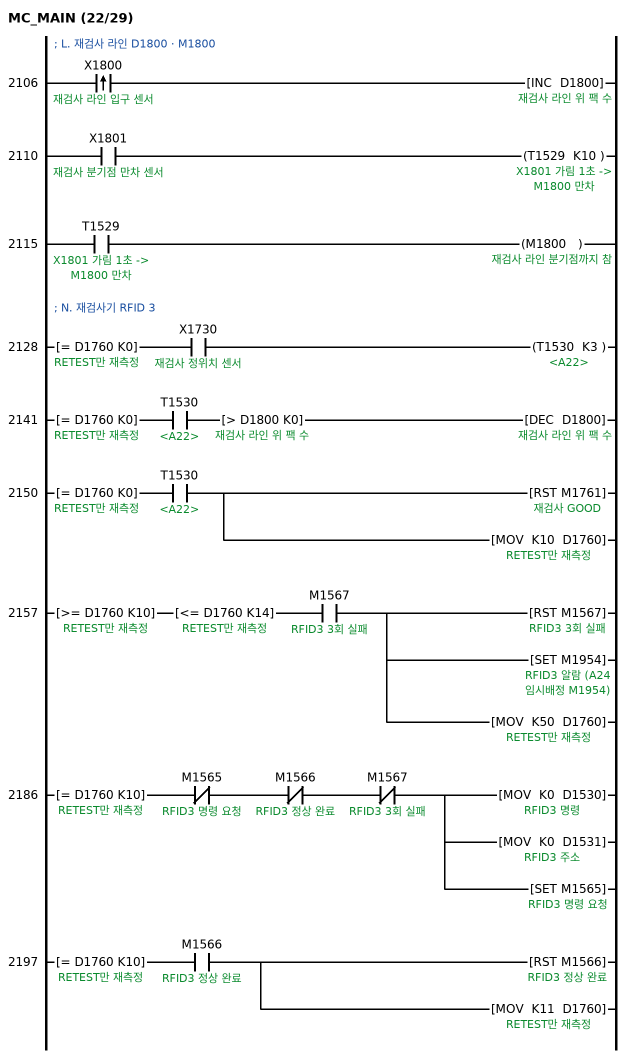
[picture p24: ladder of MC_MAIN, rungs at steps 2106 to 2197]
; L. 재검사 라인 D1800 · M1800
2106  LDP     X1800  ; 재검사 라인 입구 센서
      INC     D1800  ; 재검사 라인 위 팩 수
2110  LD      X1801  ; 재검사 분기점 만차 센서
      OUT     T1529 K10  ; X1801 가림 1초 -> M1800 만차
2115  LD      T1529  ; X1801 가림 1초 -> M1800 만차
      OUT     M1800  ; 재검사 라인 분기점까지 참
; N. 재검사기 RFID 3
2128  LD=     D1760 K0  ; RETEST만 재측정
      AND     X1730  ; 재검사 정위치 센서
      OUT     T1530 K3  ; <A22>
        [note] <A22>
2141  LD=     D1760 K0  ; RETEST만 재측정
      AND     T1530  ; <A22>
      AND>    D1800 K0  ; 재검사 라인 위 팩 수
      DEC     D1800
2150  LD=     D1760 K0  ; RETEST만 재측정
      AND     T1530  ; <A22>
      RST     M1761  ; 재검사 GOOD
      MOV     K10 D1760
2157  LD>=    D1760 K10  ; RETEST만 재측정
      AND<=   D1760 K14  ; RETEST만 재측정
      AND     M1567  ; RFID3 3회 실패
      RST     M1567  ; RFID3 3회 실패
      SET     M1954  ; RFID3 알람 (A24 임시배정 M1954)
        [note] RFID3 알람 (A24 임시배정 M1954)
      MOV     K50 D1760
2186  LD=     D1760 K10  ; RETEST만 재측정
      ANI     M1565  ; RFID3 명령 요청
      ANI     M1566  ; RFID3 정상 완료
      ANI     M1567  ; RFID3 3회 실패
      MOV     K0 D1530  ; RFID3 명령
      MOV     K0 D1531  ; RFID3 주소
      SET     M1565  ; RFID3 명령 요청
2197  LD=     D1760 K10  ; RETEST만 재측정
      AND     M1566  ; RFID3 정상 완료
      RST     M1566  ; RFID3 정상 완료
      MOV     K11 D1760
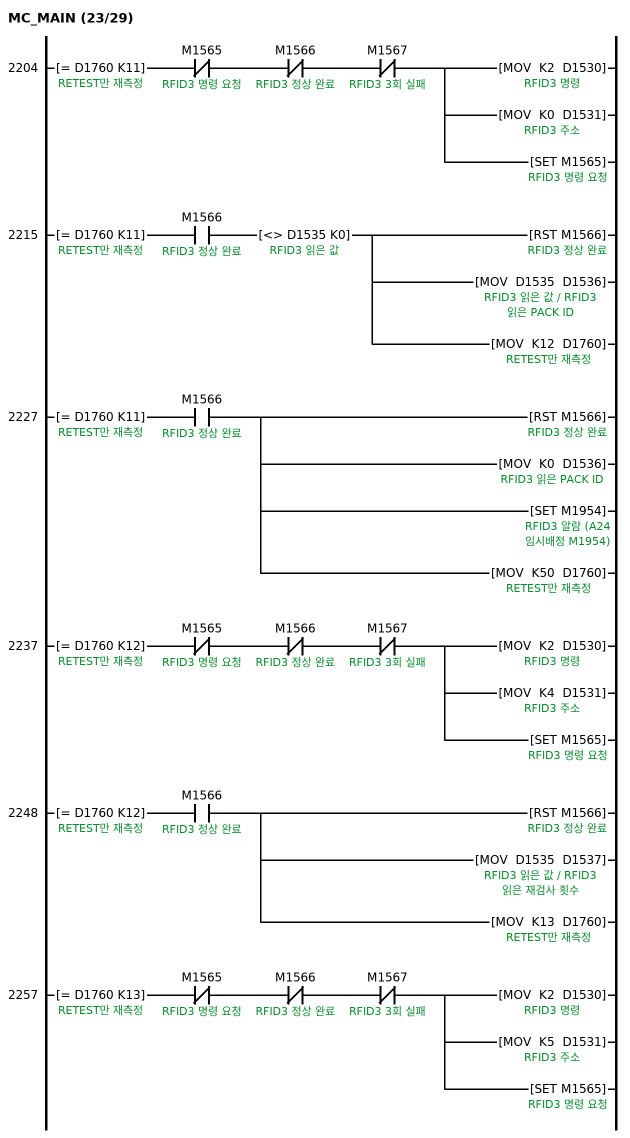
2204  LD=     D1760 K11  ; RETEST만 재측정
      ANI     M1565  ; RFID3 명령 요청
      ANI     M1566  ; RFID3 정상 완료
      ANI     M1567  ; RFID3 3회 실패
      MOV     K2 D1530
      MOV     K0 D1531
      SET     M1565  ; RFID3 명령 요청
2215  LD=     D1760 K11  ; RETEST만 재측정
      AND     M1566  ; RFID3 정상 완료
      AND<>   D1535 K0  ; RFID3 읽은 값
      RST     M1566  ; RFID3 정상 완료
      MOV     D1535 D1536  ; RFID3 읽은 PACK ID
      MOV     K12 D1760
2227  LD=     D1760 K11  ; RETEST만 재측정
      AND     M1566  ; RFID3 정상 완료
      RST     M1566  ; RFID3 정상 완료
      MOV     K0 D1536
      SET     M1954  ; RFID3 알람 (A24 임시배정 M1954)
      MOV     K50 D1760
2237  LD=     D1760 K12  ; RETEST만 재측정
      ANI     M1565  ; RFID3 명령 요청
      ANI     M1566  ; RFID3 정상 완료
      ANI     M1567  ; RFID3 3회 실패
      MOV     K2 D1530
      MOV     K4 D1531
      SET     M1565  ; RFID3 명령 요청
2248  LD=     D1760 K12  ; RETEST만 재측정
      AND     M1566  ; RFID3 정상 완료
      RST     M1566  ; RFID3 정상 완료
      MOV     D1535 D1537  ; RFID3 읽은 재검사 횟수
      MOV     K13 D1760
2257  LD=     D1760 K13  ; RETEST만 재측정
      ANI     M1565  ; RFID3 명령 요청
      ANI     M1566  ; RFID3 정상 완료
      ANI     M1567  ; RFID3 3회 실패
      MOV     K2 D1530
      MOV     K5 D1531
      SET     M1565  ; RFID3 명령 요청
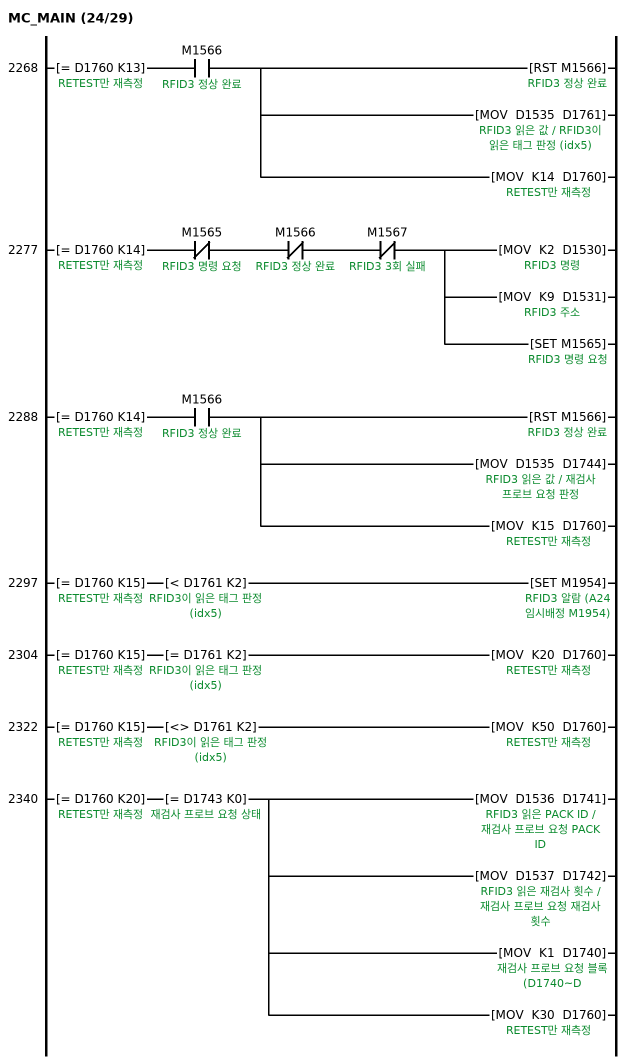
2268  LD=     D1760 K13  ; RETEST만 재측정
      AND     M1566  ; RFID3 정상 완료
      RST     M1566  ; RFID3 정상 완료
      MOV     D1535 D1761  ; RFID3이 읽은 태그 판정 (idx5)
      MOV     K14 D1760
2277  LD=     D1760 K14  ; RETEST만 재측정
      ANI     M1565  ; RFID3 명령 요청
      ANI     M1566  ; RFID3 정상 완료
      ANI     M1567  ; RFID3 3회 실패
      MOV     K2 D1530
      MOV     K9 D1531
      SET     M1565  ; RFID3 명령 요청
2288  LD=     D1760 K14  ; RETEST만 재측정
      AND     M1566  ; RFID3 정상 완료
      RST     M1566  ; RFID3 정상 완료
      MOV     D1535 D1744  ; 재검사 프로브 요청 판정
      MOV     K15 D1760
2297  LD=     D1760 K15  ; RETEST만 재측정
      AND<    D1761 K2  ; RFID3이 읽은 태그 판정 (idx5)
      SET     M1954  ; RFID3 알람 (A24 임시배정 M1954)
2304  LD=     D1760 K15  ; RETEST만 재측정
      AND=    D1761 K2  ; RFID3이 읽은 태그 판정 (idx5)
      MOV     K20 D1760
        [note] RETEST만 재측정
2322  LD=     D1760 K15  ; RETEST만 재측정
      AND<>   D1761 K2  ; RFID3이 읽은 태그 판정 (idx5)
      MOV     K50 D1760
        [note] 메인 NG -> 통과
2340  LD=     D1760 K20  ; RETEST만 재측정
      AND=    D1743 K0  ; 재검사 프로브 요청 상태
      MOV     D1536 D1741  ; 재검사 프로브 요청 PACK ID
      MOV     D1537 D1742  ; 재검사 프로브 요청 재검사 횟수
      MOV     K1 D1740  ; 재검사 프로브 요청 블록 (D1740~D
      MOV     K30 D1760
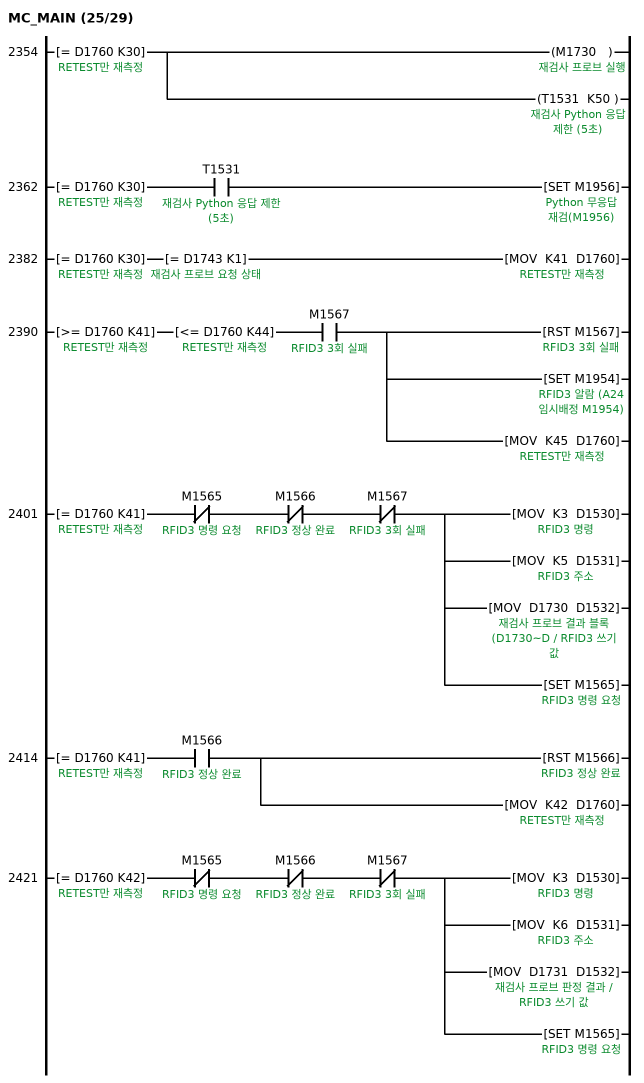
2354  LD=     D1760 K30  ; RETEST만 재측정
      OUT     M1730  ; 재검사 프로브 실행
      OUT     T1531 K50  ; 재검사 Python 응답 제한 (5초)
2362  LD=     D1760 K30  ; RETEST만 재측정
      AND     T1531  ; 재검사 Python 응답 제한 (5초)
      SET     M1956  ; Python 무응답 재검(M1956)
        [note] Python 무응답 재검(M1956)
2382  LD=     D1760 K30  ; RETEST만 재측정
      AND=    D1743 K1  ; 재검사 프로브 요청 상태
      MOV     K41 D1760
2390  LD>=    D1760 K41  ; RETEST만 재측정
      AND<=   D1760 K44  ; RETEST만 재측정
      AND     M1567  ; RFID3 3회 실패
      RST     M1567  ; RFID3 3회 실패
      SET     M1954  ; RFID3 알람 (A24 임시배정 M1954)
      MOV     K45 D1760
2401  LD=     D1760 K41  ; RETEST만 재측정
      ANI     M1565  ; RFID3 명령 요청
      ANI     M1566  ; RFID3 정상 완료
      ANI     M1567  ; RFID3 3회 실패
      MOV     K3 D1530
      MOV     K5 D1531
      MOV     D1730 D1532  ; 재검사 프로브 결과 블록 (D1730~D / RFID3 쓰기 값
      SET     M1565  ; RFID3 명령 요청
2414  LD=     D1760 K41  ; RETEST만 재측정
      AND     M1566  ; RFID3 정상 완료
      RST     M1566  ; RFID3 정상 완료
      MOV     K42 D1760
2421  LD=     D1760 K42  ; RETEST만 재측정
      ANI     M1565  ; RFID3 명령 요청
      ANI     M1566  ; RFID3 정상 완료
      ANI     M1567  ; RFID3 3회 실패
      MOV     K3 D1530
      MOV     K6 D1531
      MOV     D1731 D1532  ; 재검사 프로브 판정 결과
      SET     M1565  ; RFID3 명령 요청
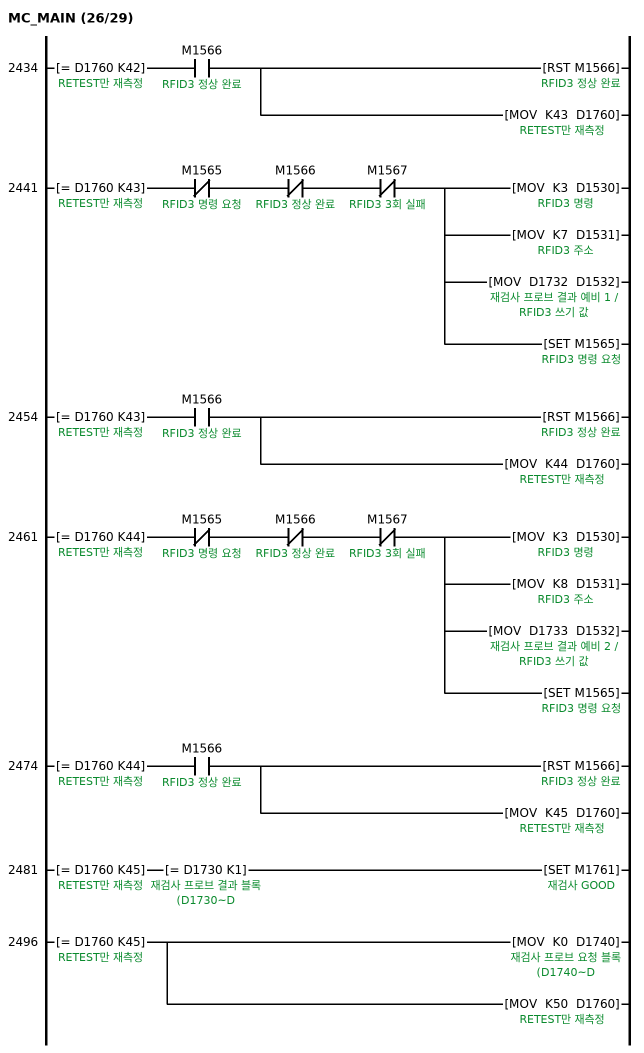
2434  LD=     D1760 K42  ; RETEST만 재측정
      AND     M1566  ; RFID3 정상 완료
      RST     M1566  ; RFID3 정상 완료
      MOV     K43 D1760
2441  LD=     D1760 K43  ; RETEST만 재측정
      ANI     M1565  ; RFID3 명령 요청
      ANI     M1566  ; RFID3 정상 완료
      ANI     M1567  ; RFID3 3회 실패
      MOV     K3 D1530
      MOV     K7 D1531
      MOV     D1732 D1532  ; 재검사 프로브 결과 예비 1
      SET     M1565  ; RFID3 명령 요청
2454  LD=     D1760 K43  ; RETEST만 재측정
      AND     M1566  ; RFID3 정상 완료
      RST     M1566  ; RFID3 정상 완료
      MOV     K44 D1760
2461  LD=     D1760 K44  ; RETEST만 재측정
      ANI     M1565  ; RFID3 명령 요청
      ANI     M1566  ; RFID3 정상 완료
      ANI     M1567  ; RFID3 3회 실패
      MOV     K3 D1530
      MOV     K8 D1531
      MOV     D1733 D1532  ; 재검사 프로브 결과 예비 2
      SET     M1565  ; RFID3 명령 요청
2474  LD=     D1760 K44  ; RETEST만 재측정
      AND     M1566  ; RFID3 정상 완료
      RST     M1566  ; RFID3 정상 완료
      MOV     K45 D1760
2481  LD=     D1760 K45  ; RETEST만 재측정
      AND=    D1730 K1  ; 재검사 프로브 결과 블록 (D1730~D
      SET     M1761  ; 재검사 GOOD
        [note] 재검사 GOOD
2496  LD=     D1760 K45  ; RETEST만 재측정
      MOV     K0 D1740
      MOV     K50 D1760
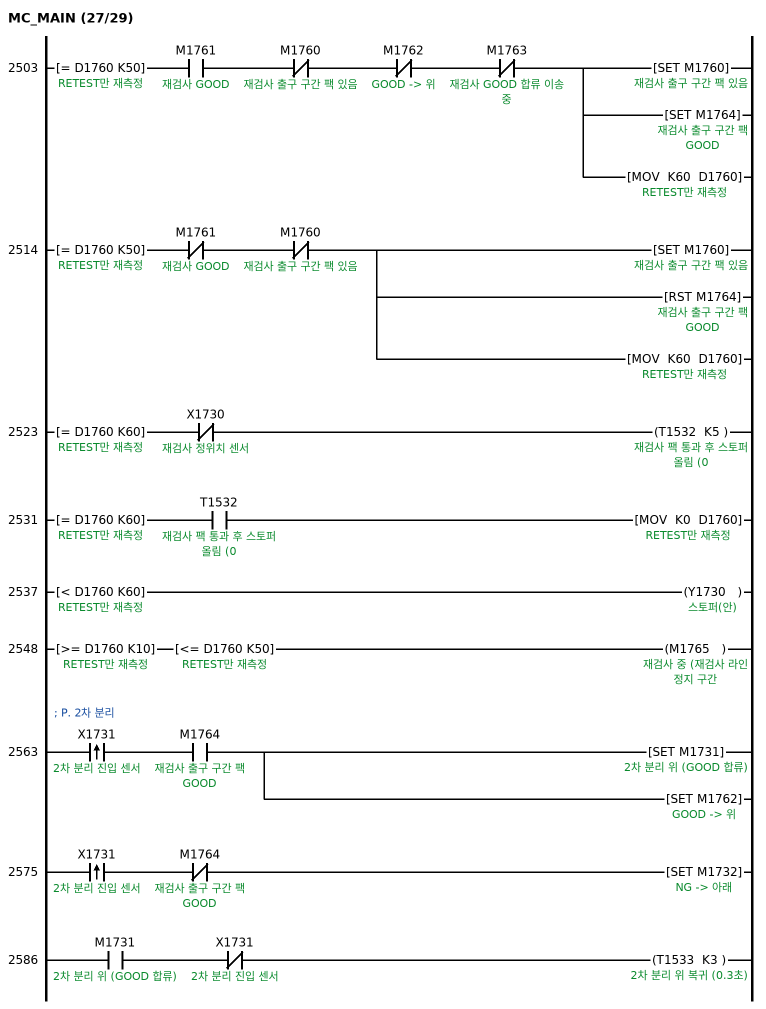
2503  LD=     D1760 K50  ; RETEST만 재측정
      AND     M1761  ; 재검사 GOOD
      ANI     M1760  ; 재검사 출구 구간 팩 있음
      ANI     M1762  ; GOOD -> 위
      ANI     M1763  ; 재검사 GOOD 합류 이송 중
      SET     M1760  ; 재검사 출구 구간 팩 있음
      SET     M1764  ; 재검사 출구 구간 팩 GOOD
      MOV     K60 D1760
2514  LD=     D1760 K50  ; RETEST만 재측정
      ANI     M1761  ; 재검사 GOOD
      ANI     M1760  ; 재검사 출구 구간 팩 있음
      SET     M1760  ; 재검사 출구 구간 팩 있음
      RST     M1764  ; 재검사 출구 구간 팩 GOOD
      MOV     K60 D1760
2523  LD=     D1760 K60  ; RETEST만 재측정
      ANI     X1730  ; 재검사 정위치 센서
      OUT     T1532 K5  ; 재검사 팩 통과 후 스토퍼 올림 (0
2531  LD=     D1760 K60  ; RETEST만 재측정
      AND     T1532  ; 재검사 팩 통과 후 스토퍼 올림 (0
      MOV     K0 D1760
2537  LD<     D1760 K60  ; RETEST만 재측정
      OUT     Y1730  ; 스토퍼(안)
        [note] 스토퍼(안)
2548  LD>=    D1760 K10  ; RETEST만 재측정
      AND<=   D1760 K50  ; RETEST만 재측정
      OUT     M1765  ; 재검사 중 (재검사 라인 정지 구간
; P. 2차 분리
2563  LDP     X1731  ; 2차 분리 진입 센서
      AND     M1764  ; 재검사 출구 구간 팩 GOOD
      SET     M1731  ; 2차 분리 위 (GOOD 합류)
      SET     M1762  ; GOOD -> 위
        [note] GOOD -> 위
2575  LDP     X1731  ; 2차 분리 진입 센서
      ANI     M1764  ; 재검사 출구 구간 팩 GOOD
      SET     M1732  ; NG -> 아래
        [note] NG -> 아래
2586  LD      M1731  ; 2차 분리 위 (GOOD 합류)
      ANI     X1731  ; 2차 분리 진입 센서
      OUT     T1533 K3  ; 2차 분리 위 복귀 (0.3초)
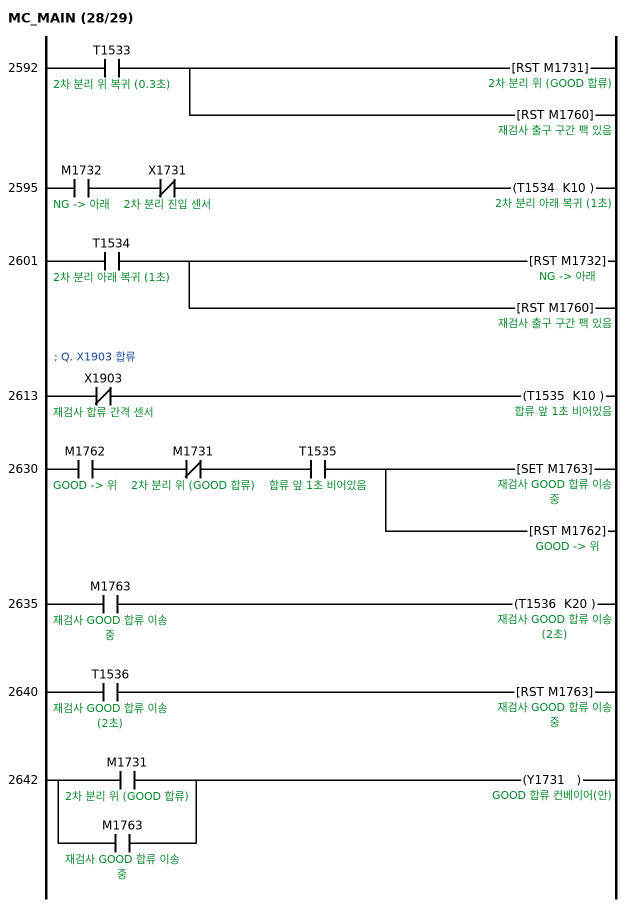
2592  LD      T1533  ; 2차 분리 위 복귀 (0.3초)
      RST     M1731  ; 2차 분리 위 (GOOD 합류)
      RST     M1760  ; 재검사 출구 구간 팩 있음
2595  LD      M1732  ; NG -> 아래
      ANI     X1731  ; 2차 분리 진입 센서
      OUT     T1534 K10  ; 2차 분리 아래 복귀 (1초)
2601  LD      T1534  ; 2차 분리 아래 복귀 (1초)
      RST     M1732  ; NG -> 아래
      RST     M1760  ; 재검사 출구 구간 팩 있음
; Q. X1903 합류
2613  LDI     X1903  ; 재검사 합류 간격 센서
      OUT     T1535 K10  ; 합류 앞 1초 비어있음
        [note] 합류 앞 1초 비어있음
2630  LD      M1762  ; GOOD -> 위
      ANI     M1731  ; 2차 분리 위 (GOOD 합류)
      AND     T1535  ; 합류 앞 1초 비어있음
      SET     M1763  ; 재검사 GOOD 합류 이송 중
      RST     M1762  ; GOOD -> 위
2635  LD      M1763  ; 재검사 GOOD 합류 이송 중
      OUT     T1536 K20  ; 재검사 GOOD 합류 이송 (2초)
2640  LD      T1536  ; 재검사 GOOD 합류 이송 (2초)
      RST     M1763  ; 재검사 GOOD 합류 이송 중
2642  LD      M1731  ; 2차 분리 위 (GOOD 합류)
      OR      M1763  ; 재검사 GOOD 합류 이송 중
      OUT     Y1731  ; GOOD 합류 컨베이어(안)
        [note] GOOD 합류 컨베이어(안)
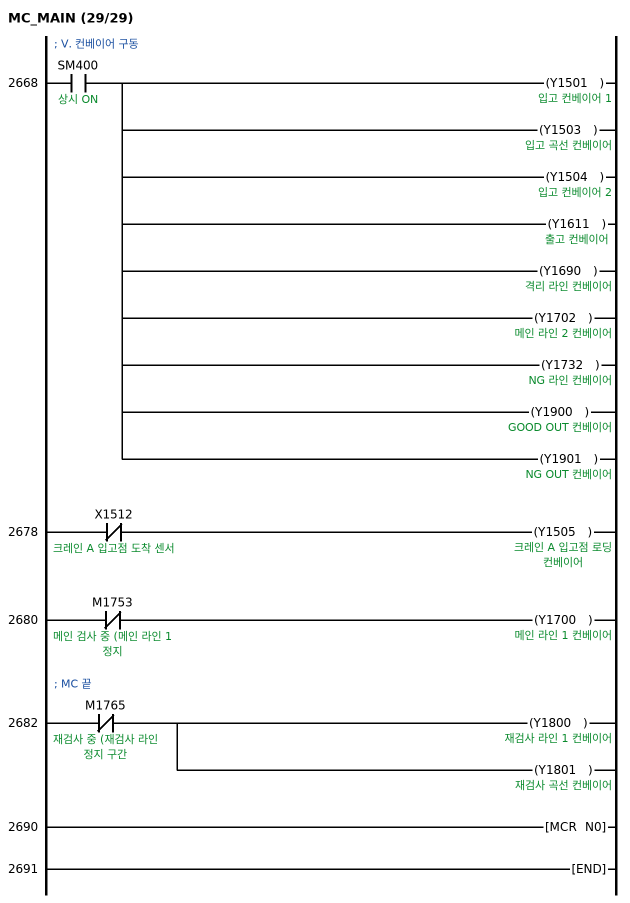
; V. 컨베이어 구동
2668  LD      SM400  ; 상시 ON
      OUT     Y1501  ; 입고 컨베이어 1
      OUT     Y1503  ; 입고 곡선 컨베이어
      OUT     Y1504  ; 입고 컨베이어 2
      OUT     Y1611  ; 출고 컨베이어
      OUT     Y1690  ; 격리 라인 컨베이어
      OUT     Y1702  ; 메인 라인 2 컨베이어
      OUT     Y1732  ; NG 라인 컨베이어
      OUT     Y1900  ; GOOD OUT 컨베이어
      OUT     Y1901  ; NG OUT 컨베이어
2678  LDI     X1512  ; 크레인 A 입고점 도착 센서
      OUT     Y1505  ; 크레인 A 입고점 로딩 컨베이어
2680  LDI     M1753  ; 메인 검사 중 (메인 라인 1 정지
      OUT     Y1700  ; 메인 라인 1 컨베이어
2682  LDI     M1765  ; 재검사 중 (재검사 라인 정지 구간
      OUT     Y1800  ; 재검사 라인 1 컨베이어
      OUT     Y1801  ; 재검사 곡선 컨베이어
; MC 끝
2690  MCR     N0
2691  END
END_PROGRAM

PROGRAM GATE_ALM
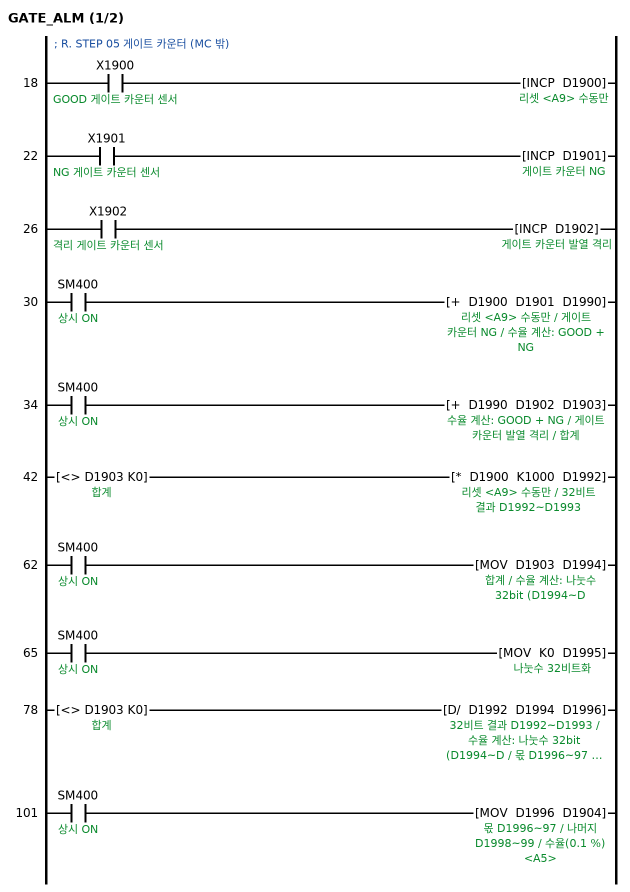
; R. STEP 05 게이트 카운터 (MC 밖)
18    LD      X1900  ; GOOD 게이트 카운터 센서
      INCP    D1900  ; 리셋 <A9> 수동만
22    LD      X1901  ; NG 게이트 카운터 센서
      INCP    D1901  ; 게이트 카운터 NG
26    LD      X1902  ; 격리 게이트 카운터 센서
      INCP    D1902  ; 게이트 카운터 발열 격리
30    LD      SM400  ; 상시 ON
      +       D1900 D1901 D1990  ; 수율 계산: GOOD + NG
34    LD      SM400  ; 상시 ON
      +       D1990 D1902 D1903  ; 합계
        [note] 합계
42    LD<>    D1903 K0  ; 합계
      *       D1900 K1000 D1992  ; 32비트 결과 D1992~D1993
        [note] 32비트 결과 D1992~D1993
62    LD      SM400  ; 상시 ON
      MOV     D1903 D1994  ; 수율 계산: 나눗수 32bit (D1994~D
65    LD      SM400  ; 상시 ON
      MOV     K0 D1995  ; 나눗수 32비트화
        [note] 나눗수 32비트화
78    LD<>    D1903 K0  ; 합계
      D/      D1992 D1994 D1996  ; 몫 D1996~97 / 나머지 D1998~99
        [note] 몫 D1996~97 / 나머지 D1998~99
101   LD      SM400  ; 상시 ON
      MOV     D1996 D1904  ; 수율(0.1 %) <A5>
        [note] 수율(0.1 %) <A5>
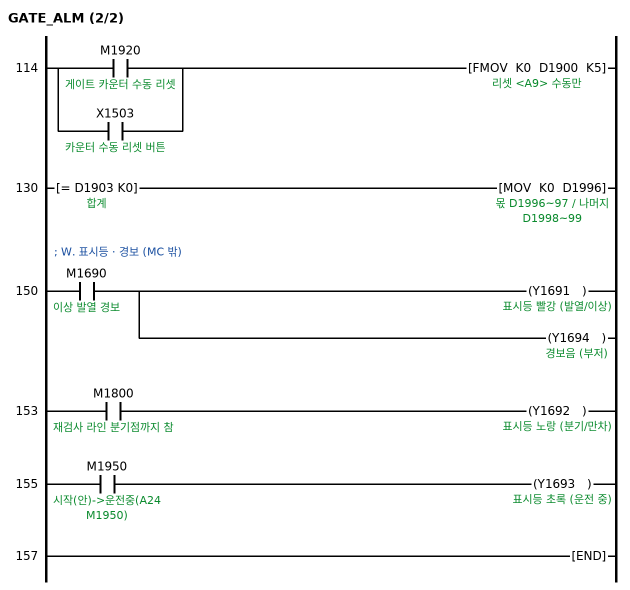
114   LD      M1920  ; 게이트 카운터 수동 리셋
      OR      X1503  ; 카운터 수동 리셋 버튼
      FMOV    K0 D1900 K5
        [note] 리셋 <A9> 수동만
130   LD=     D1903 K0  ; 합계
      MOV     K0 D1996
; W. 표시등 · 경보 (MC 밖)
150   LD      M1690  ; 이상 발열 경보
      OUT     Y1691  ; 표시등 빨강 (발열/이상)
      OUT     Y1694  ; 경보음 (부저)
153   LD      M1800  ; 재검사 라인 분기점까지 참
      OUT     Y1692  ; 표시등 노랑 (분기/만차)
155   LD      M1950  ; 시작(안)->운전중(A24 M1950)
      OUT     Y1693  ; 표시등 초록 (운전 중)
157   END
END_PROGRAM

// device comments not shown above
D1810  ; 랙 표2 칸별 입고 시각(초) R01~R2
X1511  ; 박스 높이 센서 (<A26> 1안)
X1611  ; 출고 컨베이어 센서
D1509  ; Emitter Base (<A28> 팔레트)
D1519  ; 박스 크기 판별 값 (<A26>)
D1610  ; 칸별 LOCK 경과 시간(초) R01~R24
D1660  ; 랙 표1 칸별 PACK ID R01~R24 (D16
D1840  ; 랙 표3 칸별 가상 온도/LOCK R01~R
D1870  ; 랙 표4 크레인 목표 칸 변환표 R01
